% RSLogix 500 project PROGRAM_8.RSS, saved by version 8.30.00.16 %
PROJECT "UNTITLED"    % processor: Bul.1763 MicroLogix 1100 Series B %

PROGRAM FILES
  LAD 2 "MAIN"  2 rungs
  LAD 3 "PRC_LOG"  8 rungs
  LAD 4 "OPERATIONS"  3 rungs

DATA FILES
  O0 OUTPUT  4 elements
  I1 INPUT  6 elements
  S2 STATUS  66 elements
  B3 BINARY  1 elements
  T4 TIMER  1 elements
  C5 COUNTER  1 elements
  R6 CONTROL  1 elements
  N7 INTEGER  11 elements
  F8 FLOAT  1 elements

LADDER 2 "MAIN"
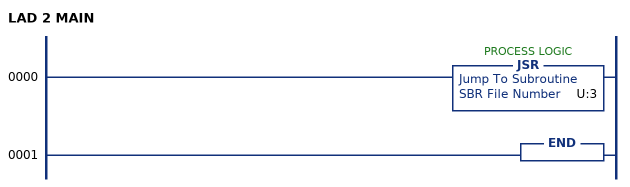
% Rung: 0 %
SOR JSR U:3 EOR
%   U:3  "PROCESS LOGIC" %
% Rung: 1 %
SOR END EOR

LADDER 3 "PRC_LOG"
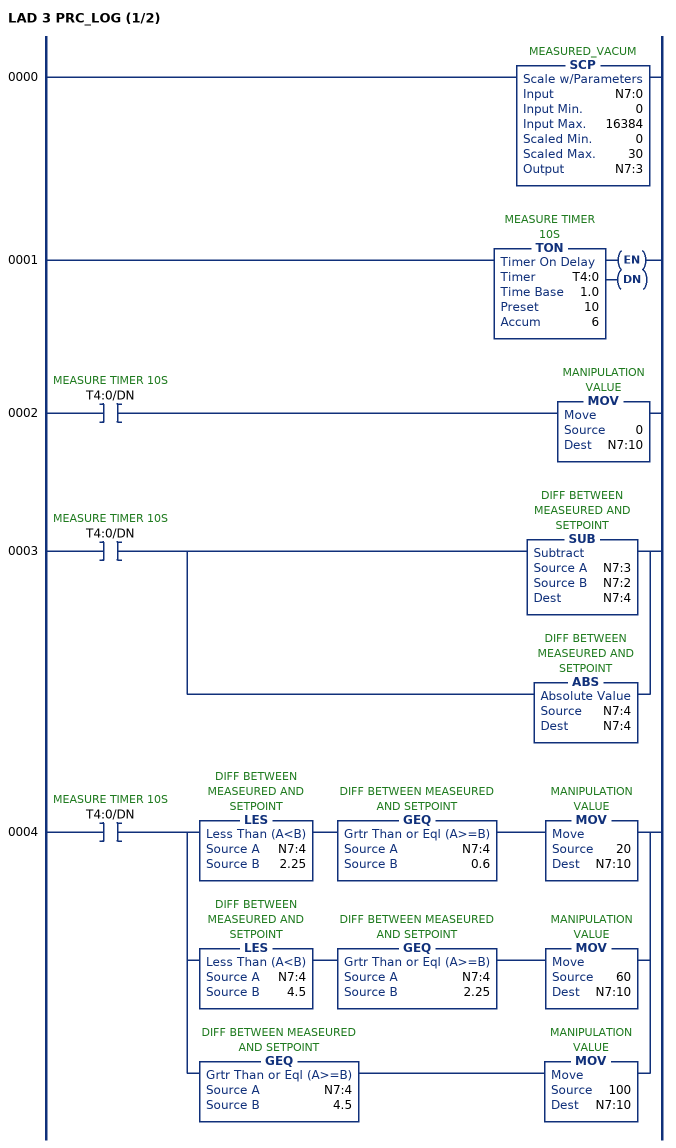
% Rung: 0 %
SOR SCP N7:0 0 16384 0 30 N7:3 EOR
%   N7:0  VACUM_SENSOR_IN %
%   N7:3  "MEASURED_VACUM" %
% Rung: 1 %
SOR TON T4:0 1.0 10 6 EOR
%   T4:0  "MEASURE TIMER 10S" %
% Rung: 2 %
SOR XIC T4:0/DN MOV 0 N7:10 EOR
%   T4:0  "MEASURE TIMER 10S" %
%   N7:10  "MANIPULATION VALUE" %
% Rung: 3 %
SOR XIC T4:0/DN BST SUB N7:3 N7:2 N7:4 NXB ABS N7:4 N7:4 BND EOR
%   T4:0  "MEASURE TIMER 10S" %
%   N7:3  "MEASURED_VACUM" %
%   N7:2  "VACUM_SETPOINT" %
%   N7:4  "DIFF BETWEEN MEASEURED AND SETPOINT" %
% Rung: 4 %
SOR XIC T4:0/DN BST LES N7:4 2.25 GEQ N7:4 0.6 MOV 20 N7:10 NXB LES N7:4 4.5 GEQ N7:4 2.25 MOV 60 N7:10 NXB GEQ N7:4 4.5 MOV 100 N7:10 BND EOR
%   T4:0  "MEASURE TIMER 10S" %
%   N7:4  "DIFF BETWEEN MEASEURED AND SETPOINT" %
%   N7:10  "MANIPULATION VALUE" %

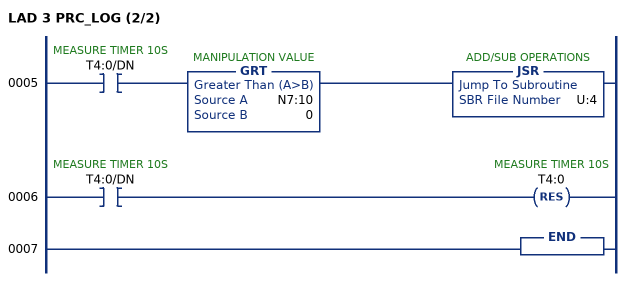
% Rung: 5 %
SOR XIC T4:0/DN GRT N7:10 0 JSR U:4 EOR
%   T4:0  "MEASURE TIMER 10S" %
%   N7:10  "MANIPULATION VALUE" %
%   U:4  "ADD/SUB OPERATIONS" %
% Rung: 6 %
SOR XIC T4:0/DN RES T4:0 EOR
%   T4:0  "MEASURE TIMER 10S" %
% Rung: 7 %
SOR END EOR

LADDER 4 "OPERATIONS"
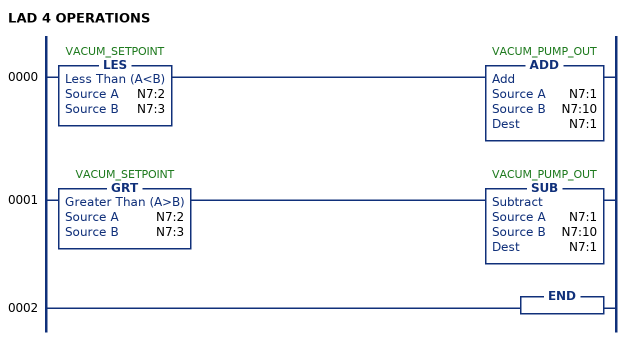
% Rung: 0 %
SOR LES N7:2 N7:3 ADD N7:1 N7:10 N7:1 EOR
%   N7:2  "VACUM_SETPOINT" %
%   N7:3  "MEASURED_VACUM" %
%   N7:1  "VACUM_PUMP_OUT" %
%   N7:10  "MANIPULATION VALUE" %
% Rung: 1 %
SOR GRT N7:2 N7:3 SUB N7:1 N7:10 N7:1 EOR
%   N7:2  "VACUM_SETPOINT" %
%   N7:3  "MEASURED_VACUM" %
%   N7:1  "VACUM_PUMP_OUT" %
%   N7:10  "MANIPULATION VALUE" %
% Rung: 2 %
SOR END EOR

OTHER DOCUMENTED ADDRESSES
  B3:0/1  "ONS"
  B3:0/2  "VACUM SENSOR BIT"
  B3:1  "ONS"
  N7:5  "DEV OF DIFFERENCE AND MEASURED POINT"
  N7:6  "ERROR VALUE"

DATA TABLE (non-zero values as saved)
DATA T4
% .PRE .ACC %
% T4:0 % 10 6
DATA N7
% N7:0 % 4000 2340 15 7 8 0 -7 0 0 0
% N7:10 % 100
DATA F8
% F8:0 % 0.0625
